(* IEC 61131-3 sources: plcassist-cli/packages/volt-lsp-iec/test-corpus/pro2193/Device/Plc Logic/Application/09 Misc/Library Manager/MemoryUtils, 6 files *)

(* ---- BITCPY.fun ---- *)
FUNCTION BITCPY : BOOL
VAR_INPUT
	PDEST : POINTER TO BYTE;
	WDSTSTARTBIT : WORD;
	PSOURCE : POINTER TO BYTE;
	WSRCSTARTBIT : WORD;
	WSIZE : WORD;
END_VAR
END_FUNCTION

(* ---- MEMCMP.fun ---- *)
FUNCTION MEMCMP : BOOL
VAR_INPUT
	PBYMEM1 : POINTER TO BYTE;
	PBYMEM2 : POINTER TO BYTE;
	DWSIZE : DWORD;
END_VAR
END_FUNCTION

(* ---- MEMFORCESWAP.fun ---- *)
FUNCTION MEMFORCESWAP : INT
VAR_INPUT
	PBYBUFFER : POINTER TO BYTE;
	ISIZE : INT;
	ICOUNT : INT;
END_VAR
END_FUNCTION

(* ---- SWAP.fun ---- *)
FUNCTION SWAP : INT
VAR_INPUT
	PUC : POINTER TO BYTE;
	ISIZE : INT;
END_VAR
END_FUNCTION

(* ---- BYTEBUFFER.fb ---- *)
FUNCTION_BLOCK BYTEBUFFER
VAR_INPUT
	PBYBUFFER : POINTER TO BYTE;
	UDIBUFFERSIZE : UDINT;
	EBYTEORDER : ByteOrder;
END_VAR
VAR_OUTPUT
	POS : UDINT;
	UDIBYTESREMAINING : UDINT;
	XOVERFLOW : BOOL;
END_VAR
VAR
	NEEDSSWAPPING : BOOL;
END_VAR
END_FUNCTION_BLOCK

METHOD ALIGN2
END_METHOD

METHOD ALIGN4
END_METHOD

METHOD CHECKOVERFLOW : BOOL
VAR_INPUT
	UDILENGTH : UDINT;
END_VAR
END_METHOD

METHOD GETBYTE : BYTE
END_METHOD

METHOD GETDWORD : DWORD
END_METHOD

METHOD GETDATAPOINTER : POINTER TO BYTE
END_METHOD

METHOD GETLWORD : LWORD
END_METHOD

METHOD GETNBYTES
VAR_INPUT
	PBYTARGET : POINTER TO BYTE;
	NBYTES : UINT;
END_VAR
END_METHOD

METHOD GETNDWORDS
VAR_INPUT
	PDWTARGET : POINTER TO DWORD;
	UICOUNT : UINT;
END_VAR
END_METHOD

METHOD GETNLWORDS
VAR_INPUT
	PDWTARGET : POINTER TO LWORD;
	UICOUNT : UINT;
END_VAR
END_METHOD

METHOD GETNWORDS
VAR_INPUT
	PWTARGET : POINTER TO WORD;
	UICOUNT : UINT;
END_VAR
END_METHOD

METHOD GETWORD : WORD
END_METHOD

METHOD INCREMENTPOS : BOOL
VAR_INPUT
	UDILENGTH : UDINT;
END_VAR
END_METHOD

METHOD PADDING
VAR_INPUT
	LEN : DINT;
END_VAR
END_METHOD

METHOD PUTBYTE
VAR_INPUT
	BYBYTE : BYTE;
END_VAR
END_METHOD

METHOD PUTDWORD
VAR_INPUT
	DWDWORD : DWORD;
END_VAR
END_METHOD

METHOD PUTLWORD
VAR_INPUT
	LWLWORD : LWORD;
END_VAR
END_METHOD

METHOD PUTNBYTES
VAR_INPUT
	PBYSOURCE : POINTER TO BYTE;
	UICOUNT : UINT;
END_VAR
END_METHOD

METHOD PUTNDWORDS
VAR_INPUT
	PDWSOURCE : POINTER TO DWORD;
	UICOUNT : UINT;
END_VAR
END_METHOD

METHOD PUTNLWORDS
VAR_INPUT
	PDWSOURCE : POINTER TO LWORD;
	UICOUNT : UINT;
END_VAR
END_METHOD

METHOD PUTNWORDS
VAR_INPUT
	PWSOURCE : POINTER TO WORD;
	UICOUNT : UINT;
END_VAR
END_METHOD

METHOD PUTWORD
VAR_INPUT
	WWORD : WORD;
END_VAR
END_METHOD

METHOD RESETPOSITION
END_METHOD

METHOD SKIP
VAR_INPUT
	LEN : UINT;
END_VAR
END_METHOD

(* ---- MEMORYMANAGER.fb ---- *)
FUNCTION_BLOCK MEMORYMANAGER
VAR
	_HXCHG : CAA.HANDLE;
	_UDIINITSIZE : UDINT;
	_UDIACTSIZE : UDINT;
	_UDIMSGLEFT : CAA.COUNT;
	_UDIBLOCKSIZE : UDINT;
	_XAUTOEXTEND : BOOL := TRUE;
	ACTSIZE : UDINT;
	AUTOEXTEND : BOOL;
	EXCHANGE : CAA.HANDLE;
	INITSIZE : UDINT;
	MESSAGESLEFT : CAA.COUNT;
END_VAR
END_FUNCTION_BLOCK

METHOD EXTEND : BOOL
VAR_INPUT
	UDINUMMSGS : UDINT;
END_VAR
END_METHOD

METHOD FB_EXIT
VAR_INPUT
	BINCOPYCODE : BOOL;
END_VAR
END_METHOD

METHOD CREATE
VAR_INPUT
	UDIINITSIZE : UDINT;
	UDIBLOCKSIZE : UDINT;
END_VAR
END_METHOD

METHOD DELETE
END_METHOD

METHOD FREE
VAR_INPUT
	PMSG : POINTER TO BYTE;
END_VAR
END_METHOD

METHOD MALLOC : POINTER TO BYTE
VAR_OUTPUT
	EERROR : ERROR;
END_VAR
END_METHOD
